FUNCTION_BLOCK F (* Negative C1: restructured by state count, returns to START every scan and dispatches on SEQ *)
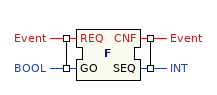
  EVENT_INPUT
    REQ WITH GO;
  END_EVENT
  EVENT_OUTPUT
    CNF WITH SEQ;
  END_EVENT
  VAR_INPUT
    GO : BOOL;
  END_VAR
  VAR_OUTPUT
    SEQ : INT;
  END_VAR
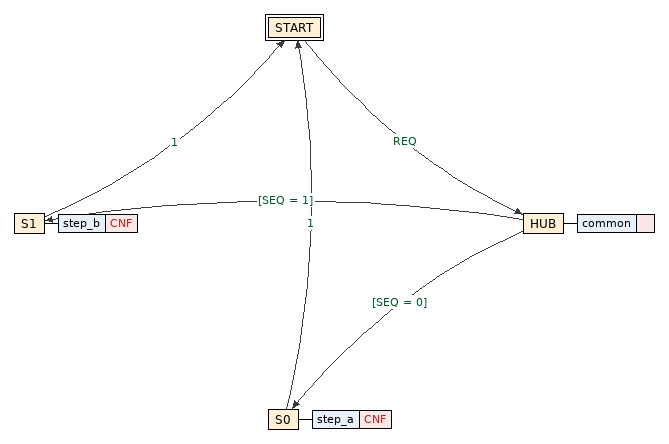
  EC_STATES
    START;
    HUB : common;
    S0 : step_a -> CNF;
    S1 : step_b -> CNF;
  END_STATES
  EC_TRANSITIONS
    START TO HUB := REQ;
    HUB TO S0 := [SEQ = 0];
    HUB TO S1 := [SEQ = 1];
    S0 TO START := 1;
    S1 TO START := 1;
  END_TRANSITIONS
  ALGORITHM common IN ST:
SEQ := SEQ;
  END_ALGORITHM
  ALGORITHM step_a IN ST:
SEQ := 0;
IF GO THEN
  SEQ := 1;
END_IF;
  END_ALGORITHM
  ALGORITHM step_b IN ST:
IF NOT GO THEN
  SEQ := 0;
END_IF;
  END_ALGORITHM
END_FUNCTION_BLOCK
